FUNCTION_BLOCK SampleFB
VAR_INPUT
	bEnable : BOOL;
END_VAR
VAR_OUTPUT
	bDone : BOOL;
END_VAR
VAR
	nCnt : INT;
END_VAR

IF bEnable THEN
	nCnt := nCnt + 1;
	bDone := nCnt >= 10;
ELSE
	nCnt := 0;
	bDone := FALSE;
END_IF

END_FUNCTION_BLOCK

(* stored: Version 1.1.0.1, ProductVersion 3.1.4024.13
   POU SampleFB: Id {aaaaaaaa-bbbb-cccc-dddd-eeeeeeeeeeee}, SpecialFunc None *)
